Fanuc KAREL source: ko00073.KL

-- PROVISIONAL review KL for V770-1; original PC SHA256 3da43b9eb950fbb1c39fd2b19ea19d1cbe854f99f71c525708f3583ea9bb0849
-- Incomplete behavior may be omitted. Consult companion uncertainty JSON. Do not deploy.
PROGRAM KO00073
%NOLOCKGROUP
BEGIN
  -- UNRESOLVED_PC offsets 5-12; opcodes 9D,23
  -- UNRESOLVED_PC offsets 17-66; opcodes 27,22,1C,27,49,7E,AD,22,31,7E,4A
  -- UNRESOLVED_PC offsets 71-75; opcodes 7F
END KO00073
